// SIMATIC S7-200 project (STEP 7-Micro/WIN), CPU 224XP CN REL 02.01

SYMBOL_TABLE USUARIO1
C_1              VD100
C_0              VD110
L_k              VD180
r_k              VD190
m_k              VD120
m_k_1            VD130
m_k_2            VD140
e_k              VD300
e_k_1            VD160
e_k_2            VD170
e_lim            VD200
h_max            VD210
Kp               VD220
h_act            VD230
Ki               VD240
r_k_1            VD250
e_ant            VD260
CONT1            VW270
CONT2            VW280
U_p              VD310
U_i_1            VD340
U_i              VD350
END_SYMBOL_TABLE

ORGANIZATION_BLOCK PRINCIPAL:OB1
TITLE=COMENTARIOS DEL PROGRAMA
BEGIN
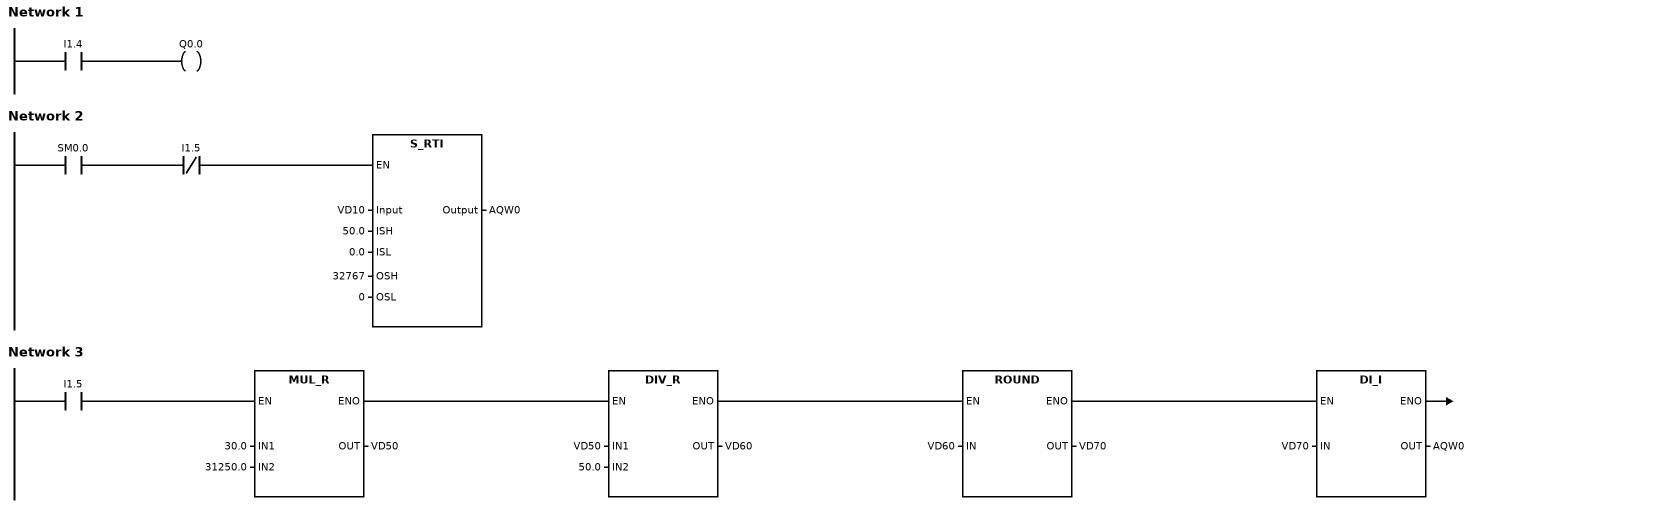
Network 1
LD     I1.4
=      Q0.0
Network 2
LD     SM0.0
AN     I1.5
CALL   S_RTI:SBR1, VD10, 50.0, 0.0, 32767, 0, AQW0
Network 3
LD     I1.5
MOVR   30.0, VD50
AENO
*R     31250.0, VD50
AENO
MOVR   VD50, VD60
AENO
/R     50.0, VD60
AENO
ROUND  VD60, VD70
AENO
DTI    VD70, AQW0
END_ORGANIZATION_BLOCK

// SBR1: protected block, not included
